{attribute 'call_after_init'}
FUNCTION_BLOCK FB_ConveyorBase
VAR_INPUT
    enable : BOOL := TRUE;
    StartDelay : TIME := T#100ms;
END_VAR
VAR_OUTPUT
    id : DINT;
    running : BOOL;
    actualSpeed : LREAL;
    ready : BOOL;
    initTrace : DINT;
    baseInitCount : DINT;
    afterInitCount : DINT;
END_VAR
VAR
    config : REFERENCE TO ST_ConveyorConfig;
    startTimer : TON;
    factor : LREAL;
END_VAR

startTimer(IN := ready AND enable AND_THEN config.enabled, PT := StartDelay);
running := startTimer.Q;
IF running THEN
    actualSpeed := config.speed * factor;
ELSE
    actualSpeed := 0.0;
END_IF;

METHOD PUBLIC FB_init : BOOL
VAR_INPUT
    bInitRetains : BOOL;
    bInCopyCode : BOOL;
    conveyorId : DINT;
    sharedConfig : REFERENCE TO ST_ConveyorConfig;
END_VAR
id := conveyorId;
config REF= sharedConfig;
baseInitCount := baseInitCount + 1;
initTrace := initTrace * 10 + 1;
FB_init := TRUE;
END_METHOD

PROPERTY PUBLIC SpeedFactor : LREAL
GET
SpeedFactor := factor;
END_GET
SET
factor := SpeedFactor;
(* Instrumentation of this example's setup order. *)
initTrace := initTrace * 10 + 3;
END_SET
END_PROPERTY

{attribute 'call_after_init'}
METHOD PUBLIC AfterInit
afterInitCount := afterInitCount + 1;
initTrace := initTrace * 10 + 4;
END_METHOD

END_FUNCTION_BLOCK

(* stored: Version 1.1.0.1, ProductVersion 3.1 *)
